(* IEC 61131-3 sources: kns-port-domestic/upstream/plc-process-lib/src/POUs/Devices/FB_ControlValve, 8 files *)

(* ---- FB_ControlValve.decl.st ---- *)
// Назначение: регулирующий клапан с позиционером 4–20 мА. Задание положения с пределами и
//             ограничением скорости (рампа, не зависящая от цикла), плотное закрытие, инверсия
//             выхода; контроль рассогласования с ОС положения (предупреждение или фиксируемый
//             отказ по конфигурации), отказ ОС, отказ позиционера; положение безопасности по
//             блокировке и отказу мимо рампы; выход xAutoActive для слежения ПИД. Режимы Auto,
//             Manual, Local (позиционер на месте — выход следит за ОС), OutOfService (удержание).
//             Наследует FB_DeviceBase: тело — нормативный порядок цикла (раздел 9.4 контракта).
// Автор:      kr0nsch
// Версия:     0.1.0
// Документ:   docs/fb/FB_ControlValve.md
FUNCTION_BLOCK FB_ControlValve EXTENDS FB_DeviceBase
VAR_INPUT
    rPosSpAuto_pct   : REAL;             // задание от автоматики (ПИД), % хода
    rPosFb_pct       : REAL;             // ОС положения, % (обычно fbZT.rValue_pct)
    xPosFbValid      : BOOL;             // ОС достоверна (обычно fbZT.xValid)
    xLocal           : BOOL;             // позиционер в местном/ручном (байпас, маховик)
    wInterlock       : WORD := 16#0000;  // блокировки: бит = 1 — в rSafePos_pct
    xPositionerFault : BOOL;             // авария позиционера (DI) или отказ канала AO (диагностика модуля)
END_VAR
VAR_IN_OUT
    stCmd    : ST_ControlValveCmd;       // команды HMI/SCADA (GVL_Hmi.st<TAG>Cmd)
    stRetain : ST_DeviceRetain;          // режим, OOS (GVL_Persist.st<TAG>Retain)
END_VAR
VAR_IN_OUT CONSTANT
    stCfg : ST_ControlValveCfg;          // параметры (GVL_Persist.st<TAG>Cfg)
END_VAR
VAR_OUTPUT
    rOut_pct    : REAL;                  // задание положения, % хода (до инверсии)
    rOut_mA     : REAL := 4.0;           // на AO с учётом инверсии, мА
    xAutoActive : BOOL;                  // клапан следует rPosSpAuto_pct — ПИД: xTrack := NOT xAutoActive
    stSts       : ST_ControlValveSts;    // состояние для HMI/SCADA
END_VAR
VAR
    stCfgLkg     : ST_ControlValveCfg;   // последняя корректная конфигурация (LKG, нормативно)
    lrRamp_pct   : LREAL;                // положение до плотного закрытия — состояние рампы, % (LREAL, CV-14)
    xTightAct    : BOOL;                 // плотное закрытие действует (с гистерезисом CV_TIGHT_HYST_PCT, CV-13)
    xRampingPrev : BOOL;                 // в прошлом вызове рампа была активна
    xDevLatched  : BOOL;                 // зафиксированный отказ рассогласования (xDevIsFault)
    wIlkPrev     : WORD;                 // блокировки после маски в прошлом вызове (первопричина)
    uiFirstOut   : UINT := GVL_Const.NO_FIRST_OUT;   // номер бита первой блокировки; NO_FIRST_OUT — нет
    fbDev        : FB_Delay;             // задержка рассогласования tDev
    // --- сигналы и условия этого вызова: считает тело, читает шаг SelectOutput ---
    lrDt_s       : LREAL;                // шаг времени, с
    xRemote      : BOOL;                 // режим Auto или Manual
    wIlk         : WORD;                 // блокировки после маски
    xIlkAct      : BOOL;                 // блокировка действует (Auto/Manual)
    xFbOk        : BOOL;                 // ОС подключена, достоверна и конечна
    xFaultAny    : BOOL;                 // есть отказ (wFault <> 0)
    // --- результат выбора выхода этого вызова (пишет SelectOutput) ---
    rSpAct       : REAL;                 // задание после пределов, до рампы, %
    xSafe        : BOOL;                 // выход принудительно в положение безопасности
    xRamping     : BOOL;                 // рампа не дошла до задания
    xLimMin      : BOOL;                 // задание ограничено снизу
    xLimMax      : BOOL;                 // задание ограничено сверху
    xSpInvalid   : BOOL;                 // задание не конечно, выход удерживается
END_VAR
VAR_TEMP
    xResetNow  : BOOL;                   // Reset в этом вызове
    eRes       : E_CmdResult;            // результат ProcessMode
    wBit       : WORD;                   // бит при поиске первопричины
    uiBit      : UINT;                   // номер бита при поиске первопричины
    xFbInvalid : BOOL;                   // ОС подключена, но недостоверна
    xPosFault  : BOOL;                   // отказ позиционера (не в OutOfService)
    xDevCond   : BOOL;                   // условие рассогласования до задержки
    xDevWarn   : BOOL;                   // рассогласование — предупреждение
    xManualCtl : BOOL;                   // выходом управляет оператор (Manual без блокировки и отказа)
    rTightOff  : REAL;                   // положение снятия плотного закрытия, %
    xInvert    : BOOL;                   // инверсия выхода мА
    wFltBits   : WORD;                   // wFault
    wWrnBits   : WORD;                   // wWarning
    wLowBits   : WORD;                   // младший байт wStatus
    eDevSt     : E_Ne107Status;          // вклад устройства в NE 107
    xAvailDev  : BOOL;                   // готовность для автоматики (без учёта Cfg)
    xAtSp      : BOOL;                   // |выход - ОС| <= rDevMax_pct
END_VAR

(* ---- CheckConfig.method.decl.st ---- *)
// Проверка конфигурации: биты wCfgErr регулирующего клапана (CV_CFG_*). Только считает, ничего не
// меняет. Неконечные значения (NaN, ±Inf) проверяются отдельно: сравнения с NaN ложны
METHOD PROTECTED CheckConfig : WORD
VAR_IN_OUT CONSTANT
    stCfgIn : ST_ControlValveCfg;   // проверяемая конфигурация
END_VAR
VAR
    wErr : WORD;                    // непройденные проверки
END_VAR

(* ---- CheckConfig.method.impl.st ---- *)
IF NOT F_IsFinite(rIn := stCfgIn.rOutMin_pct) OR NOT F_IsFinite(rIn := stCfgIn.rOutMax_pct)
   OR stCfgIn.rOutMin_pct < 0.0 OR stCfgIn.rOutMax_pct > GVL_Const.PCT_FULL
   OR stCfgIn.rOutMin_pct >= stCfgIn.rOutMax_pct
THEN
    wErr := wErr OR GVL_Const.CV_CFG_LIMITS;
END_IF
IF NOT F_IsFinite(rIn := stCfgIn.rRateUp_pctps) OR NOT F_IsFinite(rIn := stCfgIn.rRateDown_pctps)
   OR stCfgIn.rRateUp_pctps < 0.0 OR stCfgIn.rRateDown_pctps < 0.0
THEN
    wErr := wErr OR GVL_Const.CV_CFG_RATE;
END_IF
IF NOT F_IsFinite(rIn := stCfgIn.rSafePos_pct) OR stCfgIn.rSafePos_pct < 0.0
   OR stCfgIn.rSafePos_pct > GVL_Const.PCT_FULL
THEN
    wErr := wErr OR GVL_Const.CV_CFG_SAFE_POS;
END_IF
IF stCfgIn.xFbUsed AND (NOT F_IsFinite(rIn := stCfgIn.rDevMax_pct) OR stCfgIn.rDevMax_pct <= 0.0
                        OR stCfgIn.tDev <= T#0S)
THEN
    wErr := wErr OR GVL_Const.CV_CFG_DEVIATION;
END_IF
IF NOT F_IsFinite(rIn := stCfgIn.rTightShut_pct) OR stCfgIn.rTightShut_pct < 0.0
   OR stCfgIn.rTightShut_pct >= stCfgIn.rOutMax_pct
THEN
    wErr := wErr OR GVL_Const.CV_CFG_TIGHT_SHUT;
END_IF
IF stCfgIn.eFaultAction <> E_CvFaultAction.Hold AND stCfgIn.eFaultAction <> E_CvFaultAction.SafePos THEN
    wErr := wErr OR GVL_Const.CV_CFG_FAULT_ACTION;
END_IF
IF NOT CheckAlarmCfg(astCfg := stCfgIn.astAlarm) THEN
    wErr := wErr OR GVL_Const.CV_CFG_ALARM;
END_IF
CheckConfig := wErr;

(* ---- FB_ControlValve.impl.st ---- *)
// 0. Первый вызов: число слотов тревог и тип устройства (до ProcessMode)
IF xFirstCall THEN
    uiAlarmCount := GVL_Const.CV_ALARM_COUNT;
    eDevType := E_DeviceType.ControlValve;
END_IF

// 1. Время
BeginCycle();
lrDt_s := F_LTimeToSec(ltIn := ltDt);

// 2. Конфигурация (LKG)
IF AcceptCfg(wErr := CheckConfig(stCfgIn := stCfg)) THEN
    stCfgLkg := stCfg;
END_IF

// 3. Reset: снимает зафиксированное рассогласование и первопричину. Причина рассогласования —
//    расхождение выхода и ОС за время tDev: после Reset она оценивается заново, с начала отсчёта
xResetNow := xResetReq OR stCmd.stCommon.xReset;
IF xResetNow THEN
    xDevLatched := FALSE;
    uiFirstOut := GVL_Const.NO_FIRST_OUT;
    fbDev.Preset(xValue := FALSE);
    SetCmdResult(eResult := E_CmdResult.Accepted);
END_IF

// 4. Режим: регулирующий клапан не «движется» как механизм — вывод из работы всегда допустим
eRes := ProcessMode(xLocalSel := xLocal, xLocalSupported := TRUE, xOosAllowed := TRUE,
                    stCmd := stCmd.stCommon, stRetain := stRetain);
IF eRes <> E_CmdResult.None THEN
    SetCmdResult(eResult := eRes);
END_IF

// 5. Команд-импульсов у клапана нет: задание Manual — значение stCmd.rPosSpMan_pct

// 6. Логика по stCfgLkg
xRemote := eMode = E_DeviceMode.Auto OR eMode = E_DeviceMode.Manual;
wIlk := wInterlock AND stCfgLkg.wInterlockMask;
xIlkAct := xRemote AND wIlk <> 0;
// 6.1 Первопричина: при переходе слова блокировок из 0 в не 0 — номер младшего взведённого бита
IF wIlkPrev = 0 AND wIlk <> 0 AND eMode <> E_DeviceMode.OutOfService THEN
    wBit := 1;
    uiBit := 0;
    WHILE (wIlk AND wBit) = 0 DO
        wBit := SHL(wBit, 1);
        uiBit := uiBit + 1;
    END_WHILE
    uiFirstOut := uiBit;
END_IF
wIlkPrev := wIlk;

// 6.2 ОС положения и позиционер
xFbOk := stCfgLkg.xFbUsed AND xPosFbValid AND F_IsFinite(rIn := rPosFb_pct);
xFbInvalid := stCfgLkg.xFbUsed AND NOT xFbOk;
xPosFault := xPositionerFault AND eMode <> E_DeviceMode.OutOfService;

// 6.3 Рассогласование: выход прошлого вызова против ОС этого (ОС отражает уже поданное задание);
//     только в Auto/Manual, при достоверной ОС, не во время рампы и не в первом вызове (выхода ещё не было)
xDevCond := xFbOk AND xRemote AND NOT xRampingPrev AND NOT xFirstCall
            AND ABS(rOut_pct - rPosFb_pct) > stCfgLkg.rDevMax_pct;
fbDev(xIn := xDevCond, tOnDelay := stCfgLkg.tDev, itfTime := itfTimeAct);
IF fbDev.xOut AND stCfgLkg.xDevIsFault THEN
    xDevLatched := TRUE;
END_IF
xDevWarn := fbDev.xOut AND NOT stCfgLkg.xDevIsFault;
xFaultAny := xDevLatched OR xPosFault;

// 6.4 Выбор выхода по старшинству (метод SelectOutput)
SelectOutput(rManSp_pct := stCmd.rPosSpMan_pct, rCfgSafePos_pct := stCfg.rSafePos_pct);

// 6.5 Плотное закрытие с гистерезисом (CV-13): включается ниже rTightShut_pct, снимается при положении не ниже
//     rTightShut_pct + CV_TIGHT_HYST_PCT (не выше rOutMax_pct) — задание, шумящее у порога, не «стучит» клапаном о
//     седло. Затем мА с инверсией (без корректной Cfg — инверсия из поданной Cfg)
rTightOff := MIN(stCfgLkg.rTightShut_pct + GVL_Const.CV_TIGHT_HYST_PCT, stCfgLkg.rOutMax_pct);
IF stCfgLkg.rTightShut_pct <= 0.0 THEN
    xTightAct := FALSE;
ELSIF lrRamp_pct < REAL_TO_LREAL(stCfgLkg.rTightShut_pct) THEN
    xTightAct := TRUE;
ELSIF lrRamp_pct >= REAL_TO_LREAL(rTightOff) THEN
    xTightAct := FALSE;
END_IF
IF xTightAct THEN
    rOut_pct := 0.0;
ELSE
    rOut_pct := LREAL_TO_REAL(lrRamp_pct);
END_IF
IF xCfgEverOk THEN
    xInvert := stCfgLkg.xOutInvert;
ELSE
    xInvert := stCfg.xOutInvert;
END_IF
IF xInvert THEN
    rOut_mA := GVL_Const.MA_ZERO + GVL_Const.MA_SPAN * (GVL_Const.PCT_FULL - rOut_pct) / GVL_Const.PCT_FULL;
ELSE
    rOut_mA := GVL_Const.MA_ZERO + GVL_Const.MA_SPAN * rOut_pct / GVL_Const.PCT_FULL;
END_IF

// 6.6 Слежение: пока выходом управляет не оператор, задание Manual = текущий выход
xManualCtl := xCfgEverOk AND eMode = E_DeviceMode.Manual AND NOT xIlkAct AND NOT xFaultAny;
IF NOT xManualCtl THEN
    stCmd.rPosSpMan_pct := rOut_pct;
END_IF
xRampingPrev := xRamping;

// 7. Тревоги (слоты E_CvAlarm)
axAlmCond[E_CvAlarm.Deviation] := xDevWarn OR xDevLatched;
axAlmCond[E_CvAlarm.FbFailure] := xFbInvalid;
axAlmCond[E_CvAlarm.PositionerFault] := xPosFault;
axAlmCond[E_CvAlarm.InterlockAct] := xIlkAct;
arAlmValue[E_CvAlarm.Deviation] := SEL(xFbOk, 0.0, rOut_pct - rPosFb_pct);
arAlmValue[E_CvAlarm.FbFailure] := rPosFb_pct;
arAlmValue[E_CvAlarm.PositionerFault] := rOut_pct;
arAlmValue[E_CvAlarm.InterlockAct] := rOut_pct;
RunAlarms(udiIdBase := stCfgLkg.udiAlarmIdBase, stCmd := stCmd.stCommon, astCfg := stCfgLkg.astAlarm);

// 8. Состояние
xAtSp := xFbOk AND ABS(rOut_pct - rPosFb_pct) <= stCfgLkg.rDevMax_pct;
wFltBits := SEL(xDevLatched, 0, GVL_Const.CV_FLT_DEVIATION) OR SEL(xPosFault, 0, GVL_Const.CV_FLT_POSITIONER);
wWrnBits := SEL(xDevWarn, 0, GVL_Const.CV_WRN_DEVIATION)
            OR SEL(xFbInvalid, 0, GVL_Const.CV_WRN_FB_INVALID)
            OR SEL(xSpInvalid, 0, GVL_Const.CV_WRN_SP_INVALID);
xAvailDev := eMode = E_DeviceMode.Auto AND wFltBits = 0 AND wIlk = 0;
xAutoActive := xAvailDev AND xCfgEverOk;
wLowBits := SEL(xAtSp, 0, GVL_Const.CV_STS_AT_SETPOINT)
            OR SEL(xRamping, 0, GVL_Const.CV_STS_RAMPING)
            OR SEL(xLimMin, 0, GVL_Const.CV_STS_LIMITED_MIN)
            OR SEL(xLimMax, 0, GVL_Const.CV_STS_LIMITED_MAX)
            OR SEL(xIlkAct, 0, GVL_Const.CV_STS_INTERLOCKED)
            OR SEL(xTightAct, 0, GVL_Const.CV_STS_TIGHT_SHUT)
            OR SEL(xSafe, 0, GVL_Const.CV_STS_SAFE_POS)
            OR SEL(xAutoActive, 0, GVL_Const.CV_STS_AVAILABLE);
IF wFltBits <> 0 THEN
    eDevSt := E_Ne107Status.Failure;
ELSIF xDevWarn THEN
    eDevSt := E_Ne107Status.OutOfSpecification;
ELSIF xFbInvalid THEN
    eDevSt := E_Ne107Status.MaintenanceRequired;
ELSE
    eDevSt := E_Ne107Status.Good;
END_IF
stSts.rPosSp_pct := rSpAct;
stSts.rOut_pct := rOut_pct;
stSts.rOut_mA := rOut_mA;
// ОС в Sts — конечная (NaN из Modbus — 0.0, R6); достоверность — в битах
stSts.rPosFb_pct := SEL(F_IsFinite(rIn := rPosFb_pct), 0.0, rPosFb_pct);
IF xFbOk THEN
    stSts.rDeviation_pct := rOut_pct - rPosFb_pct;
ELSE
    stSts.rDeviation_pct := 0.0;
END_IF
stSts.wInterlock := wIlk;
stSts.uiFirstOut := uiFirstOut;
FinishCycle(eDevStatus := eDevSt, xAvailableDev := xAvailDev, wLow := wLowBits, wFaultBits := wFltBits,
            wWarnBits := wWrnBits, stCommon := stSts.stCommon);

(* ---- OnModeChanged.method.decl.st ---- *)
// Хук смены режима: сначала база (SUPER^); рампа предустанавливается текущим выходом (без рывка);
// вход в OutOfService снимает фиксацию рассогласования и первопричину. VAR_IN_OUT устройства не
// трогает (R2)
METHOD PROTECTED OnModeChanged
VAR_INPUT
    eOld : E_DeviceMode;   // режим до смены
    eNew : E_DeviceMode;   // новый режим
END_VAR

(* ---- OnModeChanged.method.impl.st ---- *)
SUPER^.OnModeChanged(eOld := eOld, eNew := eNew);
lrRamp_pct := REAL_TO_LREAL(rOut_pct);
IF eNew = E_DeviceMode.OutOfService THEN
    xDevLatched := FALSE;
    fbDev.Preset(xValue := FALSE);
    uiFirstOut := GVL_Const.NO_FIRST_OUT;
END_IF

(* ---- SelectOutput.method.decl.st ---- *)
// Шаг 6.4: выбор выхода по старшинству (раздел 16.3 контракта): нет корректной Cfg — положение
// безопасности из поданной Cfg; OutOfService — удержание; Local — следит за ОС (в пределах 0…100 %);
// блокировка или отказ с SafePos — rSafePos_pct мимо пределов и рампы; отказ с Hold — удержание;
// Auto/Manual — пределы и рампа (LREAL, F_RateLimitLr). lrRamp_pct — положение до плотного закрытия. Значения из
// VAR_IN_OUT — параметрами (R2).
// Шаг тела FB_ControlValve; внутренний: PROTECTED (правило L5 контракта), имя зарезервировано
METHOD PROTECTED SelectOutput
VAR_INPUT
    rManSp_pct      : REAL;   // stCmd.rPosSpMan_pct — задание оператора, %
    rCfgSafePos_pct : REAL;   // stCfg.rSafePos_pct — положение безопасности поданной Cfg, %
END_VAR
VAR
    rSpRaw    : REAL;         // задание до пределов, %
    rSafe_pct : REAL;         // положение безопасности без корректной Cfg, %
END_VAR

(* ---- SelectOutput.method.impl.st ---- *)
xSafe := FALSE;
xRamping := FALSE;
xLimMin := FALSE;
xLimMax := FALSE;
xSpInvalid := FALSE;
IF NOT xCfgEverOk THEN
    // корректной Cfg не было: положение безопасности из поданной Cfg, в 0…100; NaN — 0
    rSafe_pct := rCfgSafePos_pct;
    IF F_IsFinite(rIn := rSafe_pct) THEN
        rSpAct := LIMIT(0.0, rSafe_pct, GVL_Const.PCT_FULL);
    ELSE
        rSpAct := 0.0;
    END_IF
    lrRamp_pct := REAL_TO_LREAL(rSpAct);
    xSafe := TRUE;
ELSIF eMode = E_DeviceMode.OutOfService THEN
    rSpAct := LREAL_TO_REAL(lrRamp_pct);
ELSIF eMode = E_DeviceMode.Local THEN
    // позиционер на месте: выход следит за ОС (возврат без рывка), без ОС — удержание. ОС датчика
    // чуть выходит за 0…100 % (-1 %, 102 %) — выход в пределах хода, ток не выходит из 4…20 мА
    IF xFbOk THEN
        lrRamp_pct := REAL_TO_LREAL(LIMIT(0.0, rPosFb_pct, GVL_Const.PCT_FULL));
    END_IF
    rSpAct := LREAL_TO_REAL(lrRamp_pct);
ELSIF xIlkAct OR (xFaultAny AND stCfgLkg.eFaultAction = E_CvFaultAction.SafePos) THEN
    // блокировка и отказ с SafePos: мимо пределов и рампы — безопасность важнее плавности
    lrRamp_pct := REAL_TO_LREAL(stCfgLkg.rSafePos_pct);
    xSafe := TRUE;
    rSpAct := stCfgLkg.rSafePos_pct;
ELSIF xFaultAny THEN
    rSpAct := LREAL_TO_REAL(lrRamp_pct);
ELSE
    IF eMode = E_DeviceMode.Auto THEN
        rSpRaw := rPosSpAuto_pct;
    ELSE
        rSpRaw := rManSp_pct;
    END_IF
    IF F_IsFinite(rIn := rSpRaw) THEN
        rSpAct := LIMIT(stCfgLkg.rOutMin_pct, rSpRaw, stCfgLkg.rOutMax_pct);
        xLimMin := rSpRaw < stCfgLkg.rOutMin_pct;
        xLimMax := rSpRaw > stCfgLkg.rOutMax_pct;
        // рампа в LREAL (CV-14): приращение медленной рампы при коротком цикле не теряется округлением до REAL
        IF lrDt_s > 0.0 THEN
            lrRamp_pct := F_RateLimitLr(lrCurrent := lrRamp_pct, rTarget := rSpAct,
                                        rRateUp_ups := stCfgLkg.rRateUp_pctps,
                                        rRateDown_ups := stCfgLkg.rRateDown_pctps, lrDt_s := lrDt_s);
        ELSIF (REAL_TO_LREAL(rSpAct) > lrRamp_pct AND stCfgLkg.rRateUp_pctps <= 0.0)
              OR (REAL_TO_LREAL(rSpAct) < lrRamp_pct AND stCfgLkg.rRateDown_pctps <= 0.0)
        THEN
            // шага времени нет (первый вызов, время назад), а скорость не ограничена — сразу к заданию
            lrRamp_pct := REAL_TO_LREAL(rSpAct);
        END_IF
        xRamping := lrRamp_pct <> REAL_TO_LREAL(rSpAct);
    ELSE
        // NaN из Modbus/ПИД: удержание и предупреждение
        xSpInvalid := TRUE;
        rSpAct := LREAL_TO_REAL(lrRamp_pct);
    END_IF
END_IF
